ABB RAPID module: Feature.mod

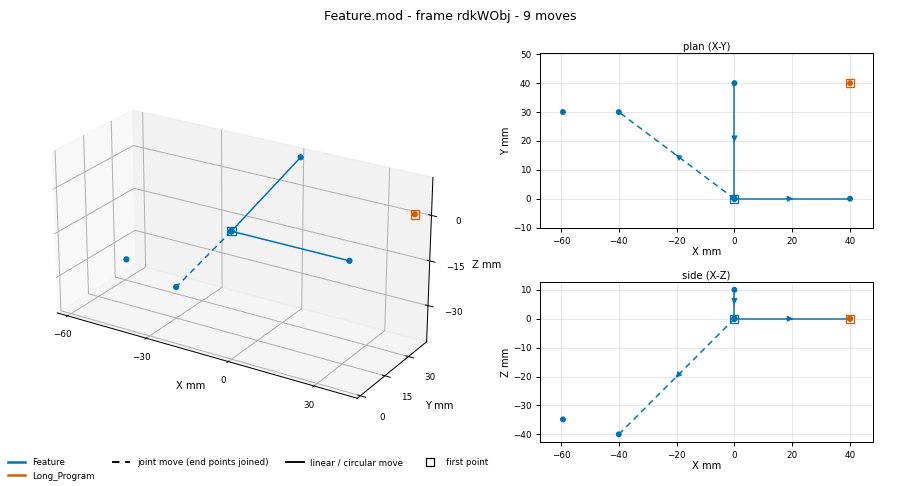
[picture p0: tool path of Feature.mod in frame rdkWObj, 9 of 13 moves have a stored position in this frame; points joined in program order, loops and branches not executed]
MODULE MOD_Feature

PERS wobjdata rdkWObj := [FALSE, TRUE, "", [[0,0,0],[1,0,0,0]],[[0,0,0],[1,0,0,0]]];
PERS tooldata rdkTool := [TRUE,[[0,0,0],[1,0,0,0]],[6.8,[0,0,15],[1,0,0,0],0,0,0.005]];
VAR speeddata rdkSpeed := [500,500,500,500];
VAR zonedata rdkZone := z1;
VAR extjoint rdkExtax := [9E9,9E9,9E9,9E9,9E9,9E9];

PROC main_RoboDK()
	Feature;
	EXIT;
ENDPROC

PROC Feature()
	!Program generated by RoboDK v5.9.4 for ABB IRB 1600-8/1.45 on 26/10/2026 01:01:07
	!Using nominal kinematics.
	var robtarget crt;
	crt := CRobT(\Tool:=rdkTool, \WObj:=rdkWObj);
	rdkExtax := crt.extax;
	ConfJ \On;
	ConfL \Off;
	rdkWObj.uframe:=[[0.000,0.000,0.000],[1.00000000,0.00000000,0.00000000,0.00000000]];
	rdkWObj.oframe:=[[851.624,-621.056,1118.740],[0.96592583,0.00000000,0.00000000,0.25881905]];
	rdkTool.tframe:=[[0.000,0.000,120.000],[0.99144486,0.00000000,0.13052619,0.00000001]];
	MoveAbsJ [[-42.973281,13.470468,-8.833703,-85.040881,-43.174179,83.214813],rdkExtax], rdkSpeed, rdkZone, rdkTool, \WObj:=rdkWObj;
	rdkSpeed:=[250.0,500,250.0,500];
	rdkZone:=z5;
	MoveJ [[0.000,0.000,0.000],[0.58801837,0.20533497,0.76632048,-0.15755906],[-1,-1,0,1],rdkExtax], rdkSpeed, rdkZone, rdkTool, \WObj:=rdkWObj;
	MoveL [[40.000,0.000,0.000],[0.58801837,0.20533497,0.76632048,-0.15755906],[-1,-1,0,1],rdkExtax], rdkSpeed, rdkZone, rdkTool, \WObj:=rdkWObj;
	MoveL CalcRobT([[-42.161283,15.522104,-11.964699,-86.080052,-42.283058,84.708364],rdkExtax], rdkTool \WObj:=rdkWObj), rdkSpeed, rdkZone, rdkTool, \WObj:=rdkWObj;
	MoveC [[40.000,40.000,0.000],[0.58801837,0.20533497,0.76632048,-0.15755906],[-1,-1,0,1],rdkExtax], [[0.000,40.000,10.000],[0.58801837,0.20533497,0.76632048,-0.15755906],[-1,-1,0,1],rdkExtax], rdkSpeed, rdkZone, rdkTool, \WObj:=rdkWObj;
	rdkZone:=fine;
	AccSet 100.0, 100.0;
	rdkSpeed:=[120.0,500,120.0,500];
	MoveL [[0.000,0.000,0.000],[0.58801837,0.20533497,0.76632048,-0.15755906],[-1,-1,0,1],rdkExtax], rdkSpeed, rdkZone, rdkTool, \WObj:=rdkWObj;
	MoveL [[0.000,0.000,0.000],[0.60644490,0.33528563,0.71902231,-0.05305707],[-1,-1,1,1],rdkExtax], rdkSpeed, rdkZone, rdkTool, \WObj:=rdkWObj;
	MoveJ [[0.000,0.000,0.000],[0.58801837,0.20533497,0.76632048,-0.15755906],[-1,-1,0,1],rdkExtax], rdkSpeed, rdkZone, rdkTool, \WObj:=rdkWObj;
	AccSet 100.0, 100.0;
	rdkSpeed:=[300.0,500,300.0,500];
	AccSet 50.0, 50.0;
	SetDO 5, 1;
	SetDO 3, 0;
	WaitDI 2, 1;
	WaitDI 4, 0, \MaxTime:=2.500;
	WaitTime \InPos, 1.500;
	STOP;
	!A comment line
	TPWrite "A message";
	SubProg;
	SpacedName;
	ExternalProg;
	Long_ProgramName12;
	AnotherLong_ExternalName;
	SetRPM700;
	Ab_c;
	custom_code(1)
	ThreadProg;
	SetDO 2, 3.5;
	rdkWObj.uframe:=[[0.000,0.000,0.000],[1.00000000,0.00000000,0.00000000,0.00000000]];
	rdkWObj.oframe:=[[891.624,-651.056,1138.740],[1.00000000,0.00000000,0.00000000,0.00000000]];
	rdkTool.tframe:=[[10.000,0.000,150.000],[1.00000000,0.00000000,0.00000000,0.00000000]];
	MoveJ [[-40.000,30.000,-40.000],[0.60876142,0.00000002,0.79335335,-0.00000002],[-1,-1,0,1],rdkExtax], rdkSpeed, rdkZone, rdkTool, \WObj:=rdkWObj;
	MoveAbsJ [[-42.973281,13.470468,-8.833703,-85.040881,-43.174179,83.214813],rdkExtax], rdkSpeed, rdkZone, rdkTool, \WObj:=rdkWObj;
	MoveL [[-59.319,30.000,-34.824],[0.60876142,0.00000002,0.79335335,-0.00000002],[-1,-1,0,1],rdkExtax], rdkSpeed, rdkZone, rdkTool, \WObj:=rdkWObj;
	rdkTool.tframe:=[[0.000,0.000,120.000],[0.99144486,0.00000000,0.13052619,0.00000001]];
	rdkWObj.uframe:=[[0.000,0.000,0.000],[1.00000000,0.00000000,0.00000000,0.00000000]];
	rdkWObj.oframe:=[[851.624,-621.056,1118.740],[0.96592583,0.00000000,0.00000000,0.25881905]];
	MoveAbsJ [[-42.973281,13.470468,-8.833703,-85.040881,-43.174179,83.214813],rdkExtax], rdkSpeed, rdkZone, rdkTool, \WObj:=rdkWObj;
ENDPROC

PROC SubProg()
	!Inside sub
ENDPROC

PROC Spaced Name()
	!Spaced body
ENDPROC

PROC Long_Program Name12()
	!Long body
	rdkTool.tframe:=[[10.000,0.000,150.000],[1.00000000,0.00000000,0.00000000,0.00000000]];
	MoveL [[40.000,40.000,0.000],[0.58801837,0.20533497,0.76632048,-0.15755906],[-1,-1,0,1],rdkExtax], rdkSpeed, rdkZone, rdkTool, \WObj:=rdkWObj;
ENDPROC

PROC ThreadProg()
	!Thread body
ENDPROC

ENDMODULE
